// Mitsubishi GX Works2 project: Ex_1   PLC: FX3G

PROGRAM MAIN
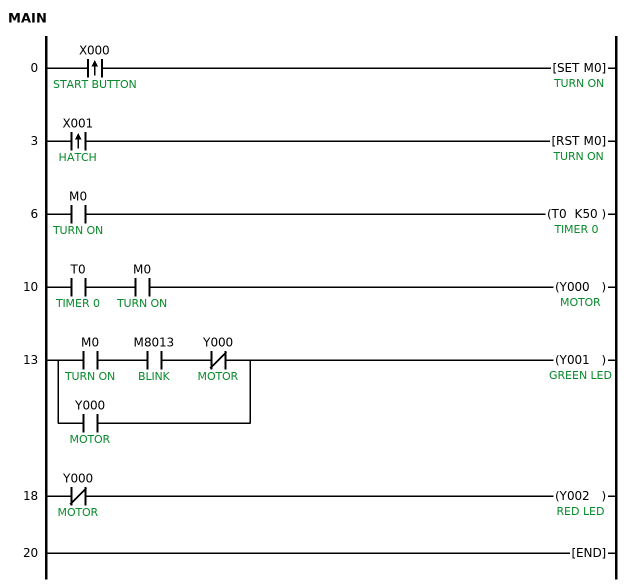
0     LDP     X000  ; START BUTTON
      SET     M0  ; TURN ON
3     LDP     X001  ; HATCH
      RST     M0  ; TURN ON
6     LD      M0  ; TURN ON
      OUT     T0 K50  ; TIMER 0
10    LD      T0  ; TIMER 0
      AND     M0  ; TURN ON
      OUT     Y000  ; MOTOR
13    LD      M0  ; TURN ON
      AND     M8013  ; BLINK
      ANI     Y000  ; MOTOR
      OR      Y000  ; MOTOR
      OUT     Y001  ; GREEN LED
18    LDI     Y000  ; MOTOR
      OUT     Y002  ; RED LED
20    END
END_PROGRAM

// device comments not shown above
T1  ; BLINK ON
T2  ; BLINK OFF
